Fanuc KAREL source: KT00902.KL

PROGRAM KT00902
%NOLOCKGROUP
VAR
  V1: VECTOR
  V2: VECTOR
  OUT: BOOLEAN
BEGIN
  V1.X = 1.0
  V2.Y = 2.0
  V1.X = 1.0
  V2.Y = 2.0
  OUT = J_IN_RANGE(V1)
END KT00902
